// TIA Portal V21 export
TextList "TL_YesNo"  ListRange=Decimal
  TextListEntry   Text="NE"
  TextListEntry   From=1, To=1, Text="DA"
